{attribute 'Tc2GvlVarNames'}
VAR_GLOBAL CONSTANT
	iSLAVEADDR_ARR_SIZE	: DINT := 256;
	dnDIAG_SLAVEINFO_SIZE	:DINT := 10;
END_VAR
VAR_GLOBAL
	SaveDiagSlaveInfo 			:ARRAY [0..dnDIAG_SLAVEINFO_SIZE] OF ST_SlaveStateInfo;
	SaveDiagSlaveInfoScanned	:ARRAY [0..dnDIAG_SLAVEINFO_SIZE] OF ST_SlaveStateInfoScanned;
END_VAR

(* stored: Version 1.1.0.1, ProductVersion 3.1.4024.15
   GVL GVL_FB_Fieldbus: Id {92384a2f-4bb3-4687-ab29-4af98505683b} *)
